// TwinCAT 3 PLC project PLC
// ProgramVersion: 3.1.4026.28
// libraries:
//   Tc2_Standard, * (Beckhoff Automation GmbH)
//   Tc2_System, * (Beckhoff Automation GmbH)
// project tree:
//   / PlcTask.TcTTO
//   POUs/ MAIN.TcPOU
// real-time tasks:
//   TASK PlcTask: cycle T#10ms, priority 20, ADS port 350

CONFIGURATION PLC
    RESOURCE PLC ON TwinCAT3
        TASK PlcTask(INTERVAL := T#10ms, PRIORITY := 20);
        PROGRAM MAIN WITH PlcTask : MAIN;
    END_RESOURCE
END_CONFIGURATION

// ---- POUs/MAIN.TcPOU
PROGRAM MAIN
VAR
	Mover  : ST_Mover;
	Active : BOOL;					// "Mover Active" - set TRUE via ADS, the PLC resets it when the arc is finished
END_VAR
VAR
	ActiveLast : BOOL;
	Angle      : LREAL;				// current angle [rad]
	AngleStep  : LREAL;				// angle increment per PLC cycle [rad]
END_VAR
VAR CONSTANT
	cPi         : LREAL := 3.14159265358979;
	cBtn        : UDINT := 1234;	// BTN the Analytics Logger condition is waiting for
	cCenterX    : LREAL := 0.0;
	cCenterY    : LREAL := 0.0;
	cRadius     : LREAL := 10.0;
	cStartAngle : LREAL := 0.0;		// Rt01 draws the first half: 0..180 deg
	cEndAngle   : LREAL := cPi;
	cArcTime    : LREAL := 5.0;		// time to draw the half circle [s]
END_VAR

Mover.ControllerID:=1; ///Who is controlling the mover - diagnostics on the scope, using dynamic sytle.

IF Active THEN
	IF NOT ActiveLast THEN
		// Rising edge: start the arc. Task cycle time is in 100 ns units.
		Angle	  := cStartAngle;
		AngleStep := (cEndAngle - cStartAngle) * UDINT_TO_LREAL(_TaskInfo[GETCURTASKINDEXEX()].CycleTime) * 1.0E-7 / cArcTime;
	END_IF

	Mover.BTN	  := cBtn;
	Mover.SetXPos := cCenterX + cRadius * COS(Angle);
	Mover.SetYPos := cCenterY + cRadius * SIN(Angle);

	IF Angle >= cEndAngle THEN
		// Finished. BTN stays 1234 for this cycle so the end point is still logged.
		Active := FALSE;
	ELSE
		Angle := MIN(Angle + AngleStep, cEndAngle);
	END_IF
ELSE
	// Inactive: only BTN drops (stops the logger). Hold the last position so the
	// one sample published after the condition clears does not spike to 0/0.
	Mover.BTN := 0;
END_IF

ActiveLast := Active;

END_PROGRAM
